(* IEC 61131-3 sources: moqui-plc/rust-plc/interfaces/codesys-system, 4 files *)

(* ---- systime.st ---- *)
(* CODESYS SysTimeRtc API used by moqui-plc. Interface declarations only (no
 * implementation). A Rust runtime maps these to the system real-time clock.
 *)

TYPE RTS_IEC_RESULT : UDINT; END_TYPE
TYPE SYSTIME : ULINT; END_TYPE

FUNCTION SysTimeRtcGet : UDINT
VAR_IN_OUT
    pResult : RTS_IEC_RESULT;
END_VAR
RETURN;
END_FUNCTION

FUNCTION SysTimeRtcConvertUtcToLocal : RTS_IEC_RESULT
VAR_INPUT
    dwTimestampUtc : UDINT;
END_VAR
VAR_IN_OUT
    pdwTimestampLocal : UDINT;
END_VAR
RETURN;
END_FUNCTION

FUNCTION SysTimeRtcHighResGet : RTS_IEC_RESULT
VAR_IN_OUT
    pTimestamp : SYSTIME;
END_VAR
RETURN;
END_FUNCTION

(* ---- device-diagnosis.st ---- *)
(* CODESYS Device Diagnosis API used by moqui-plc (library namespace DED, with
 * the CAA base types it re-exports).
 *
 * Interface declarations only (no implementation), for type checking with a
 * non-CODESYS compiler. The vendor library walks the device tree through
 * interfaces (INode, IDevice); here they are function blocks reached by
 * reference, with methods for the calls moqui-plc makes.
 *)

TYPE PVOID : POINTER TO BYTE; END_TYPE
TYPE SIZE : UDINT; END_TYPE

TYPE DED_ERROR : (NO_ERROR, INVALID_INPUT, NOT_AVAILABLE); END_TYPE
TYPE DEVICE_STATE : (UNKNOWN, NOT_CONFIGURED, OK, ERROR); END_TYPE

TYPE DEVICE_INFO :
STRUCT
    eType : DINT;
    idInstance : UDINT;
    idSystem : UDINT;
END_STRUCT
END_TYPE

FUNCTION_BLOCK INode
VAR_OUTPUT
    ChildNodeCount : UDINT;
    SiblingNodeCount : UDINT;
    FirstChildNode : REFERENCE TO INode;
    NextSiblingNode : REFERENCE TO INode;
END_VAR
END_FUNCTION_BLOCK

FUNCTION_BLOCK IDevice EXTENDS INode
VAR_OUTPUT
    Enable : BOOL;
END_VAR
METHOD GetDeviceInfo : DED_ERROR
VAR_IN_OUT
    deiInfo : DEVICE_INFO;
END_VAR
END_METHOD
METHOD GetDeviceState : DEVICE_STATE
VAR_OUTPUT
    xDiagnosisinfoAvailable : BOOL;
    eError : DED_ERROR;
END_VAR
END_METHOD
METHOD GetDeviceDiagnosisInfo : DED_ERROR
VAR_INPUT
    pData : PVOID;
    szSize : SIZE;
END_VAR
VAR_OUTPUT
    szCount : SIZE;
END_VAR
END_METHOD
END_FUNCTION_BLOCK

FUNCTION INode_TO_IDevice : REFERENCE TO IDevice
VAR_INPUT
    itfNode : REFERENCE TO INode;
END_VAR
RETURN;
END_FUNCTION

FUNCTION GetDeviceNameString : STRING
VAR_INPUT
    itfDevice : REFERENCE TO IDevice;
END_VAR
RETURN;
END_FUNCTION

(* ---- ethernet.st ---- *)
(* CODESYS Ethernet I/O driver types used by moqui-plc (library namespace
 * IODrvEthernet). Interface declarations only (no implementation).
 *)

TYPE EthernetState : (NOT_CONFIGURED, CONNECTED, DISCONNECTED, SET_IP_ERROR, ERROR); END_TYPE

(* Ethernet adapter node of the device tree. *)
FUNCTION_BLOCK IoDrvEthernet EXTENDS INode
VAR_OUTPUT
    DeviceName : STRING;
    NICName : STRING;
    Enable : BOOL;
    State : EthernetState;
END_VAR
END_FUNCTION_BLOCK

(* ---- recipes.st ---- *)
(* CODESYS Recipe Management API used by moqui-plc (library namespace
 * Recipe_Management). Interface declarations only (no implementation).
 * A Rust runtime would store recipes as files under the storage path.
 *)

FUNCTION_BLOCK RecipeManCommands
METHOD SetStoragePath : DWORD
VAR_INPUT
    stPath : STRING;
END_VAR
END_METHOD
METHOD ReloadRecipes : DWORD
VAR_INPUT
    RecipeDefinitionName : STRING;
END_VAR
END_METHOD
METHOD GetRecipeNames : DWORD
VAR_INPUT
    RecipeDefinitionName : STRING;
    pStrings : POINTER TO STRING;
    iSize : INT;
    iStartIndex : INT;
END_VAR
END_METHOD
METHOD GetRecipeCount : DINT
VAR_INPUT
    RecipeDefinitionName : STRING;
END_VAR
END_METHOD
METHOD CreateRecipe : DWORD
VAR_INPUT
    RecipeDefinitionName : STRING;
    RecipeName : STRING;
END_VAR
END_METHOD
METHOD ReadAndSaveRecipe : DWORD
VAR_INPUT
    RecipeDefinitionName : STRING;
    RecipeName : STRING;
END_VAR
END_METHOD
METHOD LoadAndWriteRecipe : DWORD
VAR_INPUT
    RecipeDefinitionName : STRING;
    RecipeName : STRING;
END_VAR
END_METHOD
METHOD DeleteRecipeFile : DWORD
VAR_INPUT
    RecipeDefinitionName : STRING;
    RecipeName : STRING;
END_VAR
END_METHOD
METHOD DeleteRecipe : DWORD
VAR_INPUT
    RecipeDefinitionName : STRING;
    RecipeName : STRING;
END_VAR
END_METHOD
METHOD ResetLastError
END_METHOD
METHOD ResetLastInfo
END_METHOD
END_FUNCTION_BLOCK
